(* IEC 61131-3 sources: 2026_Projet_YGO_ExcavatriceDragage/CODE_BACKUP/CODE_20260822_IntroductionTestCI/J_SUPERVISION/_TYPES/5_ASSISTANCE_DRAGAGE, 5 files *)

(* ---- ST_ChainDredgingAssist.st ---- *)
TYPE ST_ChainDredgingAssist :
STRUCT
    Idx101_EnableDiveSearch          : BOOL; // 1 = Assistance Plongée Armée (IHM) | 0 = Désarmée
    Idx102_EnableExtractionSequence  : BOOL; // 1 = Assistance Extraction Armée (IHM) | 0 = Désarmée
    Idx103_EnableDumpAtTremie        : BOOL; // 1 = Mode Vidage Trémie Armé (IHM) | 0 = Désarmé

    Idx201_DiveReady                 : BOOL; // 1 = Assistance Plongée Prête | 0 = Non Prête
    Idx202_DiveBusy                  : BOOL; // 1 = Séquence Plongée En Cours | 0 = Repos
    Idx203_DiveDone                  : BOOL; // 1 = Fond Confirmé | 0 = En Cours
    Idx204_DiveState                 : E_DiveSearchState; // État interne séquenceur plongée
    Idx205_DiveError                 : BOOL; // 0 = Sain | 1 = Défaut Plongée
    Idx206_DiveErrorId                : WORD; // bit0: préconditions, bit1: séquence Kobold, bit2: config seuils
    Idx207_BottomTouchConfirmed      : BOOL; // 1 = Contact Fond Confirmé (Kobold ou manuel) | 0 = Non Confirmé

    Idx301_ExtractionReady           : BOOL; // 1 = Assistance Extraction Prête | 0 = Non Prête
    Idx302_ExtractionBusy            : BOOL; // 1 = Séquence Extraction En Cours | 0 = Repos
    Idx303_ExtractionDone            : BOOL; // 1 = Extraction Terminée | 0 = En Cours
    Idx304_ExtractionState           : E_ExtractionSequenceState; // État interne séquenceur extraction
    Idx305_ExtractionError           : BOOL; // 0 = Sain | 1 = Défaut Extraction
    Idx306_ExtractionErrorId          : WORD; // bit0: fond absent, bit1: fermeture, bit2: contrôle remontée, bit3: config

    Idx401_OperatorActionId          : WORD;       // Identifiant consigne opérateur conduite (0 = aucune)
    Idx402_OperatorAction            : STRING(120); // Texte consigne opérateur (secours affichage)

    Idx501_DumpAtTremieArmed         : BOOL; // 1 = Bit IHM TglEnableDumpAtTremie actif | 0 = Désarmé
    Idx502_DumpAtTremieAssistActive  : BOOL; // 1 = Mode réellement actif (armé ET Mode MAINT_N1/N2) | 0 = Inactif
    Idx503_DumpAtTremieAtTremie      : BOOL; // 1 = M3 à la position Trémie | 0 = Ailleurs
    Idx504_DumpAtTremieBucketOpenArmed : BOOL; // 1 = Ouverture benne armée par ce mode | 0 = Non armée
    Idx505_DumpAtTremieDescentLocked : BOOL; // 1 = Descente M1/M2 verrouillée (M3 hors P1/Maintenance) | 0 = Libre

    Idx601_BypassDiveActive          : BOOL; // 1 = Bypass séquence DiveSearch armé (IHM)
    Idx602_BypassKoboldBottomTouched : BOOL; // 1 = Fond confirmé par le bypass (front montant Kobold en descente)
END_STRUCT
END_TYPE

(* ---- ST_DredgingAssistCfg.st ---- *)
(* ═══════════════════════════════════════════════════════════════
   ST_DredgingAssistCfg — Réglages persistants assistants prélèvement
   📄 Doc : DOC/AF/AF_Partie-04_Mode_SemiAuto_Sequenceur_v2.1.md §3ter
   ═══════════════════════════════════════════════════════════════ *)
TYPE ST_DredgingAssistCfg :
STRUCT
    DiveStartMin_M              : REAL := 1.0;  (* Position mini M1/M2 avant plongée *)
    ImmersionUpper_M            : REAL := 0.5;  (* Borne haute fenêtre front immersion *)
    ImmersionLower_M            : REAL := -0.5; (* Borne basse fenêtre front immersion *)
    ExtractionControlDistance_M : REAL := 2.0;  (* Remontée palier 1 avant accélération *)
    TglEnableDiveSearch         : BOOL := FALSE; (* Mode assistance plongée mémorisé *)
    TglEnableExtractionSequence : BOOL := FALSE; (* Mode assistance extraction mémorisé *)
    TglEnableDumpAtTremie       : BOOL := FALSE; (* Mode assistance vidage trémie mémorisé *)
    Initialized                 : BOOL := FALSE; (* Pont persistance/IHM initialisé *)
END_STRUCT
END_TYPE

(* ---- ST_DredgingAssistCmd.st ---- *)
(* ═══════════════════════════════════════════════════════════════
   🎮 ST_DredgingAssistCmd — Sélections IHM assistance prélèvement
   ═══════════════════════════════════════════════════════════════ *)
TYPE ST_DredgingAssistCmd :
STRUCT
    TglEnableDiveSearch         : BOOL := FALSE; (* Assistance plongée active *)
    TglEnableExtractionSequence : BOOL := FALSE; (* Assistance extraction active *)
    TglBucketAtBottomConfirmed  : BOOL := FALSE; (* Attestation manuelle temporaire du fond *)
    // Bypass simplifié de la séquence FB_DiveSearch complète (préconditions
    // strictes -- benne ouverte, DiveStartMin_M, fenêtre immersion). Si TRUE, un front MONTANT
    // Kobold pendant une descente confirme directement le fond, sans passer par l'état-machine
    // FB_DiveSearch (qui continue de tourner en parallèle, inchangée -- utile pour
    // KoboldMeasureEnable). Défaut FALSE : comportement identique à avant (séquence complète
    // seule source de confirmation).
    TglBypassDiveSearchSequence : BOOL := FALSE;
    TglEnableDumpAtTremie       : BOOL := FALSE; (* : mode vidage à la trémie —
                                                     verrouille descente treuils (P1/Maintenance
                                                     uniquement) + translation M3 (proche du haut
                                                     uniquement) ; TRUE par défaut —
                                                     ⚠️ contrairement aux deux autres, ce mode
                                                     RESTREINT des mouvements existants dès le boot *)
END_STRUCT
END_TYPE

(* ---- ST_DredgingAssistHMI.st ---- *)
(* ═══════════════════════════════════════════════════════════════
   🪨 ST_DredgingAssistHMI — Échange IHM assistants prélèvement
   ═══════════════════════════════════════════════════════════════ *)
TYPE ST_DredgingAssistHMI :
STRUCT
    Cmd   : ST_DredgingAssistCmd;
    Cfg   : ST_DredgingAssistCfg;
    State : ST_DredgingAssistState;
END_STRUCT
END_TYPE

(* ---- ST_DredgingAssistState.st ---- *)
(* ═══════════════════════════════════════════════════════════════
   🚦 ST_DredgingAssistState — États publics assistance prélèvement
   ═══════════════════════════════════════════════════════════════ *)
TYPE ST_DredgingAssistState :
STRUCT
    DiveReady                  : BOOL;
    DiveBusy                   : BOOL;
    DiveDone                   : BOOL;
    DiveError                  : BOOL;
    DiveErrorId                : WORD;
    DiveState                  : E_DiveSearchState;
    BottomTouchConfirmed       : BOOL;
    ExtractionReady            : BOOL;
    ExtractionBusy             : BOOL;
    ExtractionDone             : BOOL;
    ExtractionError            : BOOL;
    ExtractionErrorId          : WORD;
    ExtractionState            : E_ExtractionSequenceState;
    OperatorActionId           : WORD;       (* Une seule consigne conduite, arbitré en PRG_09 *)
    OperatorAction             : STRING(120); (* Texte de secours ; IHM peut mapper l'identifiant *)
    // : mode vidage à la trémie (pas de FB dédié, logique combinatoire PRG_04)
    DumpAtTremieArmed          : BOOL; (* TglEnableDumpAtTremie (bit IHM brut) *)
    DumpAtTremieAssistActive   : BOOL; (* Armé ET Mode MAINT_N1/N2 (mode réellement actif) *)
    DumpAtTremieAtTremie       : BOOL; (* M3_AtTremieStable *)
    DumpAtTremieBucketOpenArmed: BOOL; (* CmdOpen_IHM déclenché par ce mode *)
    DumpAtTremieDescentLocked  : BOOL; (* DescendPermit M1/M2 forcé par ce mode (hors P1/Maintenance) *)
    // Diagnostic bypass séquence DiveSearch
    BypassDiveActive           : BOOL; (* TglBypassDiveSearchSequence armé (descente couplée en cours) *)
    BypassKoboldBottomTouched  : BOOL; (* Fond confirmé par le bypass (front montant Kobold en descente) *)
END_STRUCT
END_TYPE
